PROGRAM main
  VAR
    START AT %QX0.0 : BOOL := FALSE;
    STOP AT %QX0.1 : BOOL := FALSE;
    SYSTEM_RUN AT %QX1.0 : BOOL := FALSE;
    MOTOR AT %QX1.2 : BOOL := FALSE;
    WARNING_LIGHT AT %QX1.1 : BOOL := FALSE;
    STARTUP_TIMER : TON;
    LINE_READY : BOOL := FALSE;
    PRODUCT_SENSOR AT %QX2.0 : BOOL := FALSE;
    PROCESS_ACTIVE : BOOL := FALSE;
    PROCESS_DONE : BOOL := FALSE;
    PROCESS_TIMER : TON;
    PROCESSOR AT %QX1.3 : BOOL := FALSE;
    WAIT_CLEAR : BOOL := FALSE;
    INSPECTION_ACTIVE AT %QX1.4 : BOOL := FALSE;
    INSPECTION_DONE : BOOL := FALSE;
    INSPECTION_TIMER : TON;
    QUALITY_FAIL AT %QX2.1 : BOOL := FALSE;
    REJECT_ACTIVE AT %QX1.5 : BOOL := FALSE;
    REJECT_PULSE : BOOL := FALSE;
    PRODUCT_ACCEPTED : BOOL := FALSE;
    PRODUCT_REJECTED : BOOL := FALSE;
    REJECT_TIMER : TP;
    ACCEPT_COUNTER : CTU;
    REJECT_COUNTER : CTU;
    ACCEPT_COUNT AT %QW3 : INT := 0;
    REJECT_COUNT AT %QW4 : INT := 0;
    RESET_COUNTS AT %QX0.2 : BOOL := FALSE;
    TOTAL_PROCESSED AT %QW5 : INT := 0;
    ORDER_QUANTITY AT %QW0 : INT := 20;
    ORDER_REMAINING AT %QW6 : INT := 20;
    QUANTITY_REACHED : BOOL := FALSE;
    ORDER_COMPLETE AT %QX1.7 : BOOL := FALSE;
    BATCH_COUNTER : CTU;
    PACKAGE_COUNTER : CTU;
    PACKAGING_TIMER : TON;
    BATCH_CAPACITY AT %QW1 : INT := 10;
    BATCH_COUNT AT %QW7 : INT := 0;
    PACKAGE_COUNT AT %QW8 : INT := 0;
    BATCH_FULL : BOOL := FALSE;
    BATCH_NOT_READY : BOOL := FALSE;
    PACKAGING_ACTIVE AT %QX1.6 : BOOL := FALSE;
    PACKAGING_DONE : BOOL := FALSE;
    SIMULATOR : PRODUCT_SIMULATOR;
    DEFECT_PERCENT AT %QW2 : INT := 25;
  END_VAR

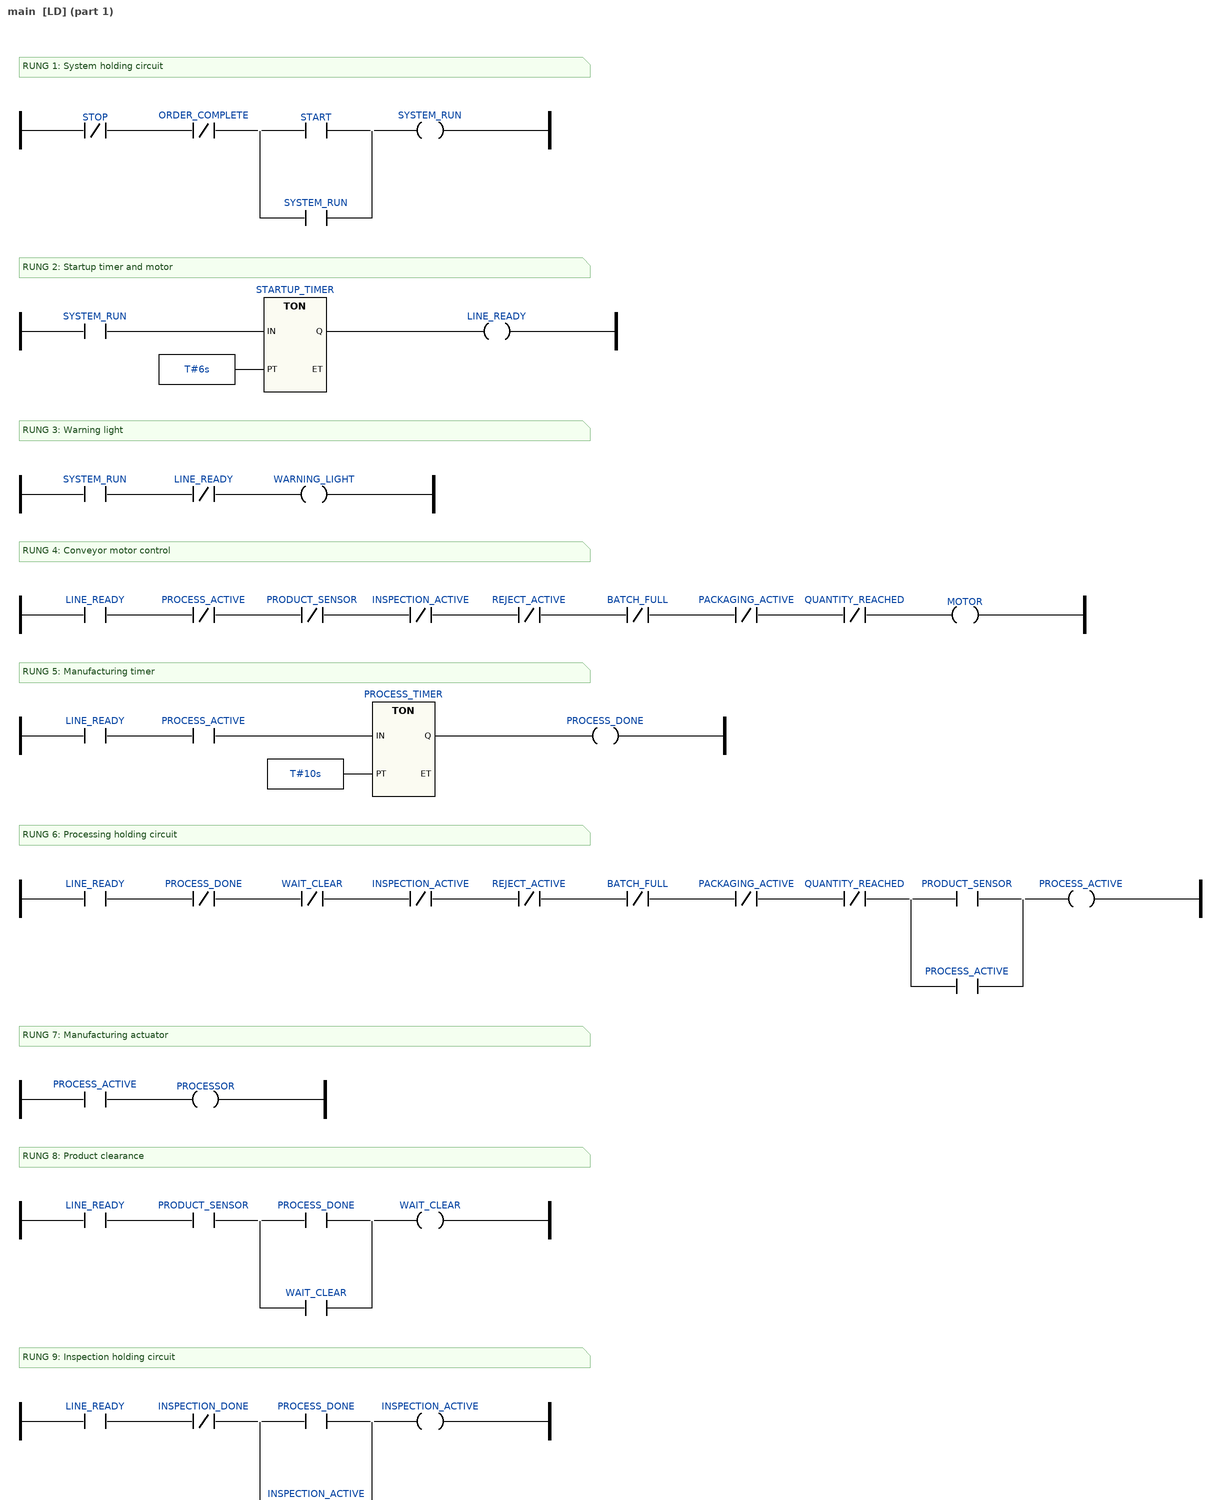
(* LD diagram, written out as Structured Text *)
(* RUNG 1: System holding circuit *)
SYSTEM_RUN := NOT STOP AND NOT ORDER_COMPLETE AND (START OR SYSTEM_RUN);
(* RUNG 2: Startup timer and motor *)
STARTUP_TIMER(IN := SYSTEM_RUN, PT := T#6s);
LINE_READY := STARTUP_TIMER.Q;
(* RUNG 3: Warning light *)
WARNING_LIGHT := SYSTEM_RUN AND NOT LINE_READY;
(* RUNG 4: Conveyor motor control *)
MOTOR := LINE_READY AND NOT PROCESS_ACTIVE AND NOT PRODUCT_SENSOR AND NOT INSPECTION_ACTIVE AND NOT REJECT_ACTIVE AND NOT BATCH_FULL AND NOT PACKAGING_ACTIVE AND NOT QUANTITY_REACHED;
(* RUNG 5: Manufacturing timer *)
PROCESS_TIMER(IN := LINE_READY AND PROCESS_ACTIVE, PT := T#10s);
PROCESS_DONE := PROCESS_TIMER.Q;
(* RUNG 6: Processing holding circuit *)
PROCESS_ACTIVE := LINE_READY AND NOT PROCESS_DONE AND NOT WAIT_CLEAR AND NOT INSPECTION_ACTIVE AND NOT REJECT_ACTIVE AND NOT BATCH_FULL AND NOT PACKAGING_ACTIVE AND NOT QUANTITY_REACHED AND (PRODUCT_SENSOR OR PROCESS_ACTIVE);
(* RUNG 7: Manufacturing actuator *)
PROCESSOR := PROCESS_ACTIVE;
(* RUNG 8: Product clearance *)
WAIT_CLEAR := LINE_READY AND PRODUCT_SENSOR AND (PROCESS_DONE OR WAIT_CLEAR);
(* RUNG 9: Inspection holding circuit *)
INSPECTION_ACTIVE := LINE_READY AND NOT INSPECTION_DONE AND (PROCESS_DONE OR INSPECTION_ACTIVE);
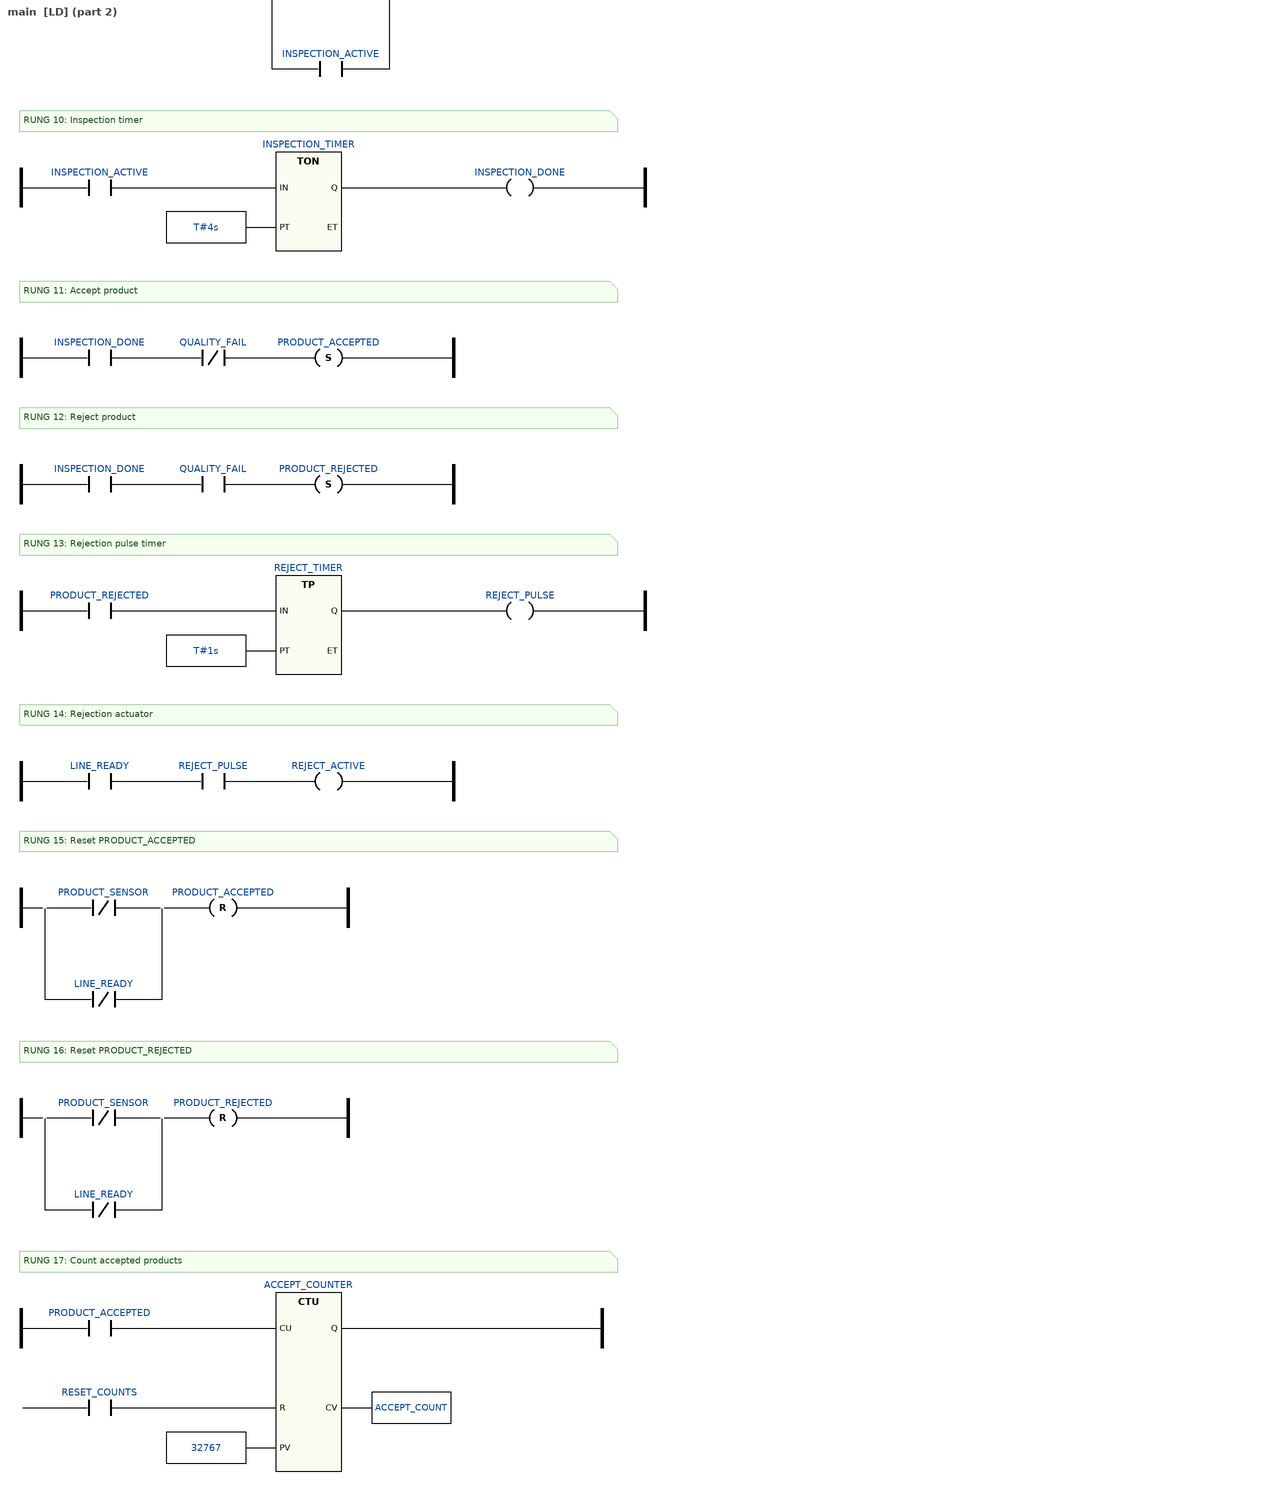
(* RUNG 10: Inspection timer *)
INSPECTION_TIMER(IN := INSPECTION_ACTIVE, PT := T#4s);
INSPECTION_DONE := INSPECTION_TIMER.Q;
(* RUNG 11: Accept product *)
IF INSPECTION_DONE AND NOT QUALITY_FAIL THEN PRODUCT_ACCEPTED := TRUE; END_IF;
(* RUNG 12: Reject product *)
IF INSPECTION_DONE AND QUALITY_FAIL THEN PRODUCT_REJECTED := TRUE; END_IF;
(* RUNG 13: Rejection pulse timer *)
REJECT_TIMER(IN := PRODUCT_REJECTED, PT := T#1s);
REJECT_PULSE := REJECT_TIMER.Q;
(* RUNG 14: Rejection actuator *)
REJECT_ACTIVE := LINE_READY AND REJECT_PULSE;
(* RUNG 15: Reset PRODUCT_ACCEPTED *)
IF NOT PRODUCT_SENSOR OR NOT LINE_READY THEN PRODUCT_ACCEPTED := FALSE; END_IF;
(* RUNG 16: Reset PRODUCT_REJECTED *)
IF NOT PRODUCT_SENSOR OR NOT LINE_READY THEN PRODUCT_REJECTED := FALSE; END_IF;
(* RUNG 17: Count accepted products *)
ACCEPT_COUNTER(CU := PRODUCT_ACCEPTED, R := RESET_COUNTS, PV := 32767);
ACCEPT_COUNT := ACCEPT_COUNTER.CV;
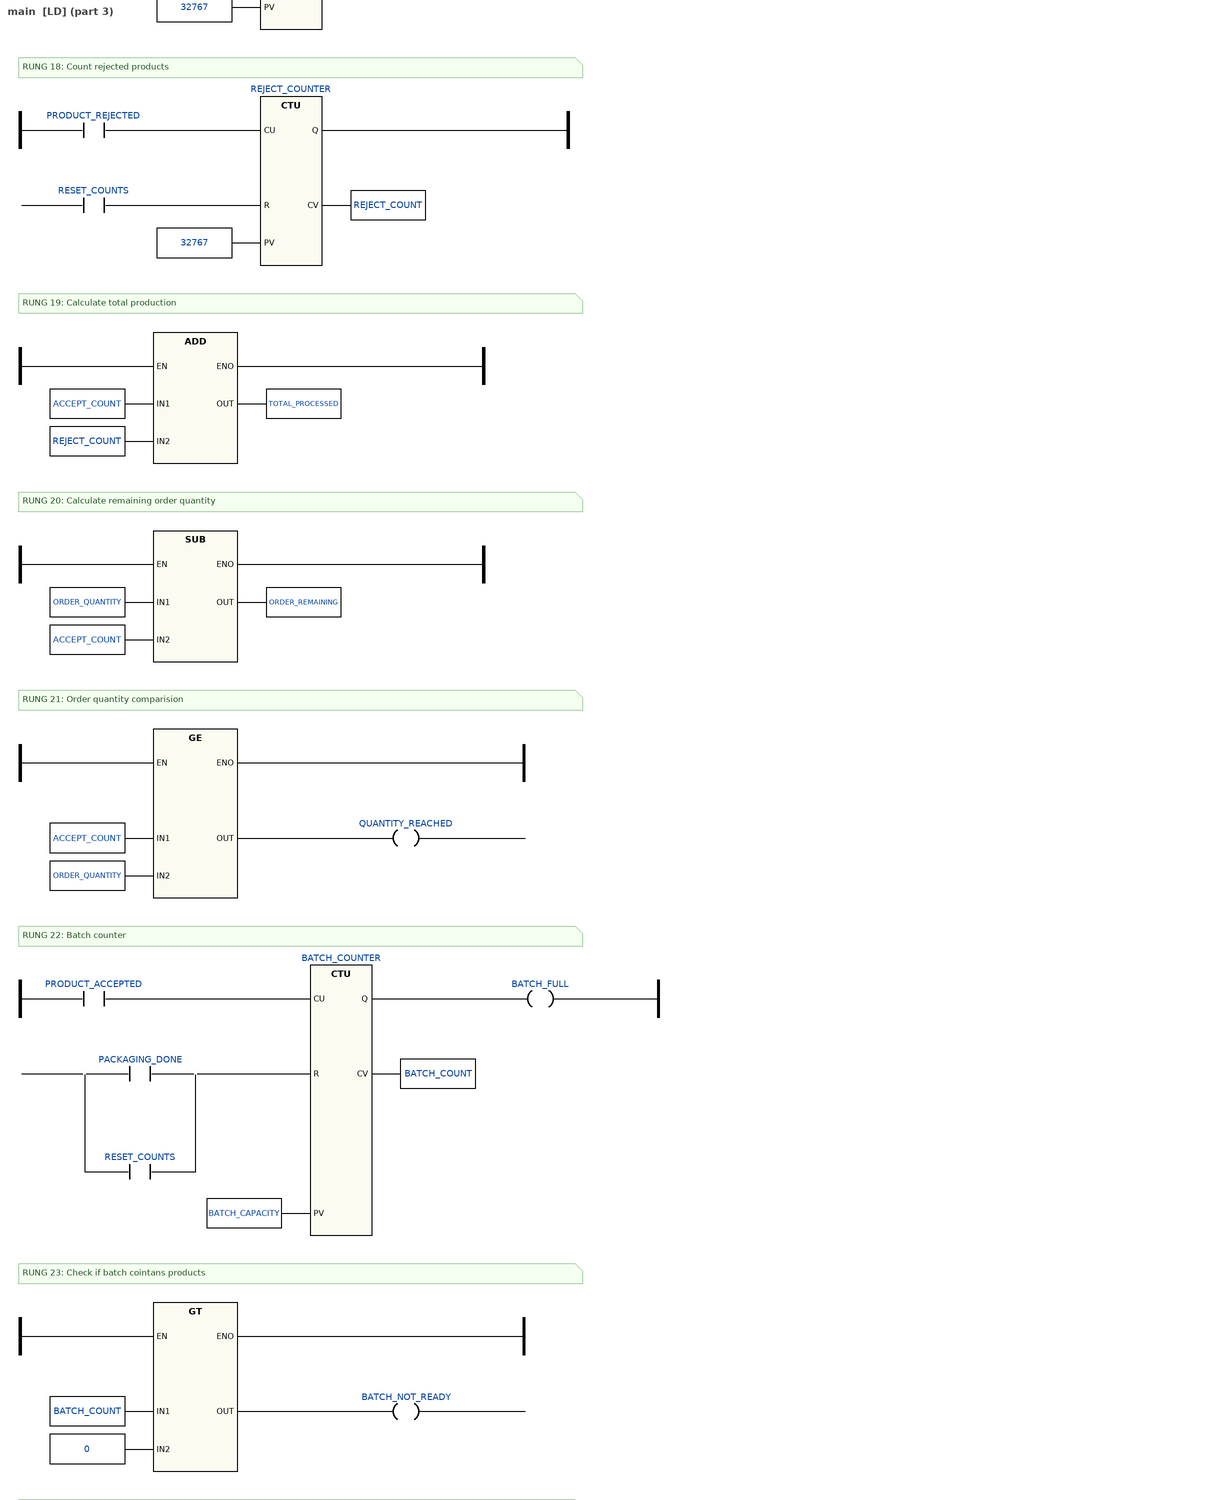
(* RUNG 18: Count rejected products *)
REJECT_COUNTER(CU := PRODUCT_REJECTED, R := RESET_COUNTS, PV := 32767);
REJECT_COUNT := REJECT_COUNTER.CV;
(* RUNG 19: Calculate total production *)
TOTAL_PROCESSED := ACCEPT_COUNT + REJECT_COUNT;
(* RUNG 20: Calculate remaining order quantity *)
ORDER_REMAINING := ORDER_QUANTITY - ACCEPT_COUNT;
(* RUNG 21: Order quantity comparision *)
QUANTITY_REACHED := ACCEPT_COUNT >= ORDER_QUANTITY;
(* RUNG 22: Batch counter *)
BATCH_COUNTER(CU := PRODUCT_ACCEPTED, R := PACKAGING_DONE OR RESET_COUNTS, PV := BATCH_CAPACITY);
BATCH_FULL := BATCH_COUNTER.Q;
BATCH_COUNT := BATCH_COUNTER.CV;
(* RUNG 23: Check if batch cointans products *)
BATCH_NOT_READY := BATCH_COUNT > 0;
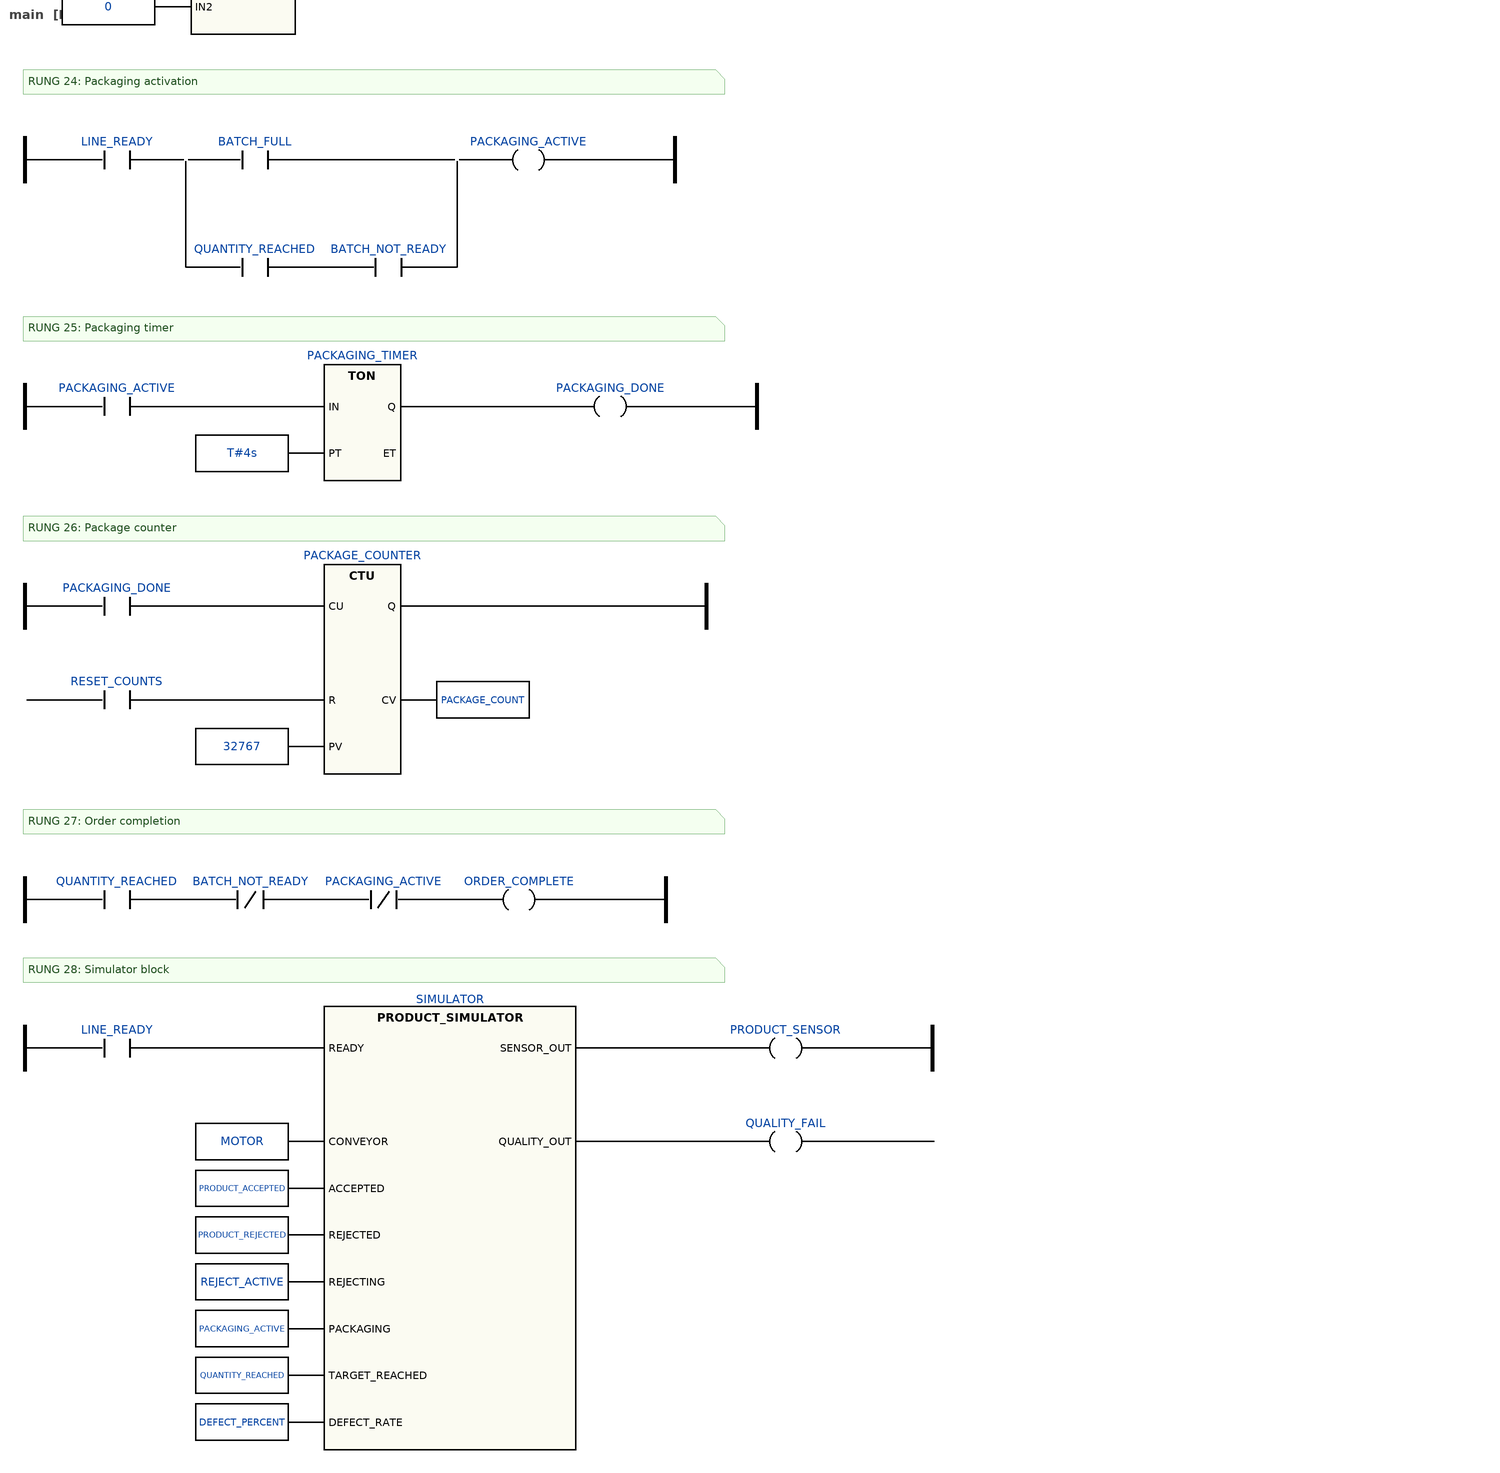
(* RUNG 24: Packaging activation *)
PACKAGING_ACTIVE := LINE_READY AND (BATCH_FULL OR QUANTITY_REACHED AND BATCH_NOT_READY);
(* RUNG 25: Packaging timer *)
PACKAGING_TIMER(IN := PACKAGING_ACTIVE, PT := T#4s);
PACKAGING_DONE := PACKAGING_TIMER.Q;
(* RUNG 26: Package counter *)
PACKAGE_COUNTER(CU := PACKAGING_DONE, R := RESET_COUNTS, PV := 32767);
PACKAGE_COUNT := PACKAGE_COUNTER.CV;
(* RUNG 27: Order completion *)
ORDER_COMPLETE := QUANTITY_REACHED AND NOT BATCH_NOT_READY AND NOT PACKAGING_ACTIVE;
(* RUNG 28: Simulator block *)
SIMULATOR(READY := LINE_READY, CONVEYOR := MOTOR, ACCEPTED := PRODUCT_ACCEPTED, REJECTED := PRODUCT_REJECTED, REJECTING := REJECT_ACTIVE, PACKAGING := PACKAGING_ACTIVE, TARGET_REACHED := QUANTITY_REACHED, DEFECT_RATE := DEFECT_PERCENT);
PRODUCT_SENSOR := SIMULATOR.SENSOR_OUT;
QUALITY_FAIL := SIMULATOR.QUALITY_OUT;
END_PROGRAM
